PROGRAM P_IEC61850_MAIN
VAR
	fbIEC 	: FB_IEC61850;	
END_VAR

fbIEC();

END_PROGRAM

(* stored: Version 1.1.0.1
   POU P_IEC61850_MAIN: Id {de4ea64a-4a85-48ba-b89c-2a3d98124197}, SpecialFunc None *)
